(* IEC 61131-3 sources: 2026_Projet_YGO_ExcavatriceDragage/CODE_BACKUP/CODE_20260904_AvantWeekendBackup_v0.6.34/J_SUPERVISION/_BRIDGES, 13 files *)

(* ---- FB_CfgPersistBridge_BucketCfg.st ---- *)
(* =======================================================================
   💾 FB_CfgPersistBridge_BucketCfg — Pont persistance pour ST_BucketCfg
   ───────────────────────────────────────────────────────────────
   🎯 Rôle : Restauration et synchronisation bidirectionnelle IHM / Persist
   💾 Persistance : Transfert GVL_PERSISTENT <-> GVL_IHM sur Initialized
   📄 Doc métier : DOC/AF/AF_Partie-03_Contrats_Composants_v2.3.md §3
   ======================================================================= *)
FUNCTION_BLOCK FB_CfgPersistBridge_BucketCfg
VAR_OUTPUT
    // === ETATS RESTAURATION ===
    JustRestored            : BOOL;               // <-- [STAT] Vrai sur le cycle de restauration initiale
END_VAR
VAR_IN_OUT
    // === BUS CONFIGURATION ET PERSISTANCE ===
    Hmi                     : ST_BucketCfg;       // <-> [BUS] Structure de configuration IHM
    Persist                 : ST_BucketCfg;       // <-> [BUS] Structure de configuration persistante
END_VAR

JustRestored := FALSE;
IF NOT Hmi.Initialized THEN
    Hmi := Persist;
    Hmi.Initialized := TRUE;
    JustRestored := TRUE;
ELSE
    Persist := Hmi;
END_IF;

(* ---- FB_CfgPersistBridge_CommunCfg.st ---- *)
(* =======================================================================
   💾 FB_CfgPersistBridge_CommunCfg — Pont persistance pour ST_CommunCfg
   ───────────────────────────────────────────────────────────────
   🎯 Rôle : Restauration et synchronisation bidirectionnelle IHM / Persist
   💾 Persistance : Transfert GVL_PERSISTENT <-> GVL_IHM sur Initialized
   📄 Doc métier : DOC/AF/AF_Partie-03_Contrats_Composants_v2.3.md §3
   ======================================================================= *)
FUNCTION_BLOCK FB_CfgPersistBridge_CommunCfg
VAR_OUTPUT
    // === ETATS RESTAURATION ===
    JustRestored            : BOOL;               // <-- [STAT] Vrai sur le cycle de restauration initiale
END_VAR
VAR_IN_OUT
    // === BUS CONFIGURATION ET PERSISTANCE ===
    Hmi                     : ST_CommunCfg;       // <-> [BUS] Structure de configuration IHM
    Persist                 : ST_CommunCfg;       // <-> [BUS] Structure de configuration persistante
END_VAR

JustRestored := FALSE;
IF NOT Hmi.Initialized THEN
    Hmi := Persist;
    Hmi.Initialized := TRUE;
    JustRestored := TRUE;
ELSE
    Persist := Hmi;
END_IF;

(* ---- FB_CfgPersistBridge_CycleAssistToggles.st ---- *)
(* =======================================================================
   💾 FB_CfgPersistBridge_CycleAssistToggles — Pont persistance toggles assistance
   ───────────────────────────────────────────────────────────────
   🎯 Rôle : Restauration et synchronisation bidirectionnelle IHM / Persist
   💾 Persistance : Transfert GVL_PERSISTENT <-> GVL_IHM sur Initialized
   📄 Doc métier : DOC/AF/AF_Partie-03_Contrats_Composants_v2.3.md §3
   ======================================================================= *)
FUNCTION_BLOCK FB_CfgPersistBridge_CycleAssistToggles
VAR_OUTPUT
    // === ETATS RESTAURATION ===
    JustRestored            : BOOL;               // <-- [STAT] Vrai sur le cycle de restauration initiale
END_VAR
VAR_IN_OUT
    // === BUS CONFIGURATION ET PERSISTANCE ===
    Hmi                     : ST_CycleAssistToggles; // <-> [BUS] Structure de toggles IHM
    Persist                 : ST_CycleAssistToggles; // <-> [BUS] Structure de toggles persistante
END_VAR

JustRestored := FALSE;
IF NOT Hmi.Initialized THEN
    Hmi := Persist;
    Hmi.Initialized := TRUE;
    JustRestored := TRUE;
ELSE
    Persist := Hmi;
END_IF;

(* ---- FB_CfgPersistBridge_CycleCfg.st ---- *)
(* =======================================================================
   💾 FB_CfgPersistBridge_CycleCfg — Pont persistance pour ST_CycleCfg
   ───────────────────────────────────────────────────────────────
   🎯 Rôle : Restauration et synchronisation bidirectionnelle IHM / Persist
   💾 Persistance : Transfert GVL_PERSISTENT <-> GVL_IHM sur Initialized
   📄 Doc métier : DOC/AF/AF_Partie-03_Contrats_Composants_v2.3.md §3
   ======================================================================= *)
FUNCTION_BLOCK FB_CfgPersistBridge_CycleCfg
VAR_OUTPUT
    // === ETATS RESTAURATION ===
    JustRestored            : BOOL;               // <-- [STAT] Vrai sur le cycle de restauration initiale
END_VAR
VAR_IN_OUT
    // === BUS CONFIGURATION ET PERSISTANCE ===
    Hmi                     : ST_CycleCfg;        // <-> [BUS] Structure de configuration IHM
    Persist                 : ST_CycleCfg;        // <-> [BUS] Structure de configuration persistante
END_VAR

JustRestored := FALSE;
IF NOT Hmi.Initialized THEN
    Hmi := Persist;
    Hmi.Initialized := TRUE;
    JustRestored := TRUE;
ELSE
    Persist := Hmi;
END_IF;

(* ---- FB_CfgPersistBridge_CycleDiveSearchCfg.st ---- *)
(* =======================================================================
   💾 FB_CfgPersistBridge_CycleDiveSearchCfg — Pont persistance cycle plongée
   ───────────────────────────────────────────────────────────────
   🎯 Rôle : Restauration et synchronisation bidirectionnelle IHM / Persist
   💾 Persistance : Transfert GVL_PERSISTENT <-> GVL_IHM sur Initialized
   📄 Doc métier : DOC/AF/AF_Partie-03_Contrats_Composants_v2.3.md §3
   ======================================================================= *)
FUNCTION_BLOCK FB_CfgPersistBridge_CycleDiveSearchCfg
VAR_OUTPUT
    // === ETATS RESTAURATION ===
    JustRestored            : BOOL;               // <-- [STAT] Vrai sur le cycle de restauration initiale
END_VAR
VAR_IN_OUT
    // === BUS CONFIGURATION ET PERSISTANCE ===
    Hmi                     : ST_CycleDiveSearchCfg; // <-> [BUS] Structure de configuration IHM
    Persist                 : ST_CycleDiveSearchCfg; // <-> [BUS] Structure de configuration persistante
END_VAR

JustRestored := FALSE;
IF NOT Hmi.Initialized THEN
    Hmi := Persist;
    Hmi.Initialized := TRUE;
    JustRestored := TRUE;
ELSE
    Persist := Hmi;
END_IF;

(* ---- FB_CfgPersistBridge_CycleDumpAtTremieCfg.st ---- *)
(* =======================================================================
   💾 FB_CfgPersistBridge_CycleDumpAtTremieCfg — Pont persistance cycle vidage trémie
   ───────────────────────────────────────────────────────────────
   🎯 Rôle : Restauration et synchronisation bidirectionnelle IHM / Persist
   💾 Persistance : Transfert GVL_PERSISTENT <-> GVL_IHM sur Initialized
   📄 Doc métier : DOC/AF/AF_Partie-03_Contrats_Composants_v2.3.md §3
   ======================================================================= *)
FUNCTION_BLOCK FB_CfgPersistBridge_CycleDumpAtTremieCfg
VAR_OUTPUT
    // === ETATS RESTAURATION ===
    JustRestored            : BOOL;               // <-- [STAT] Vrai sur le cycle de restauration initiale
END_VAR
VAR_IN_OUT
    // === BUS CONFIGURATION ET PERSISTANCE ===
    Hmi                     : ST_CycleDumpAtTremieCfg; // <-> [BUS] Structure de configuration IHM
    Persist                 : ST_CycleDumpAtTremieCfg; // <-> [BUS] Structure de configuration persistante
END_VAR

JustRestored := FALSE;
IF NOT Hmi.Initialized THEN
    Hmi := Persist;
    Hmi.Initialized := TRUE;
    JustRestored := TRUE;
ELSE
    Persist := Hmi;
END_IF;

(* ---- FB_CfgPersistBridge_CycleExtractionCfg.st ---- *)
(* =======================================================================
   💾 FB_CfgPersistBridge_CycleExtractionCfg — Pont persistance cycle extraction
   ───────────────────────────────────────────────────────────────
   🎯 Rôle : Restauration et synchronisation bidirectionnelle IHM / Persist
   💾 Persistance : Transfert GVL_PERSISTENT <-> GVL_IHM sur Initialized
   📄 Doc métier : DOC/AF/AF_Partie-03_Contrats_Composants_v2.3.md §3
   ======================================================================= *)
FUNCTION_BLOCK FB_CfgPersistBridge_CycleExtractionCfg
VAR_OUTPUT
    // === ETATS RESTAURATION ===
    JustRestored            : BOOL;               // <-- [STAT] Vrai sur le cycle de restauration initiale
END_VAR
VAR_IN_OUT
    // === BUS CONFIGURATION ET PERSISTANCE ===
    Hmi                     : ST_CycleExtractionCfg; // <-> [BUS] Structure de configuration IHM
    Persist                 : ST_CycleExtractionCfg; // <-> [BUS] Structure de configuration persistante
END_VAR

JustRestored := FALSE;
IF NOT Hmi.Initialized THEN
    Hmi := Persist;
    Hmi.Initialized := TRUE;
    JustRestored := TRUE;
ELSE
    Persist := Hmi;
END_IF;

(* ---- FB_CfgPersistBridge_CycleMachineHomingCfg.st ---- *)
(* =======================================================================
   💾 FB_CfgPersistBridge_CycleMachineHomingCfg — Pont persistance pour ST_CycleMachineHomingCfg
   ───────────────────────────────────────────────────────────────
   🎯 Rôle : Restauration et synchronisation bidirectionnelle IHM / Persist
   💾 Persistance : Transfert GVL_PERSISTENT <-> GVL_IHM sur Initialized
   📄 Doc métier : DOC/AF/AF_Partie-03_Contrats_Composants_v2.3.md §3
   ======================================================================= *)
FUNCTION_BLOCK FB_CfgPersistBridge_CycleMachineHomingCfg
VAR_OUTPUT
    // === ETATS RESTAURATION ===
    JustRestored            : BOOL;                     // <-- [STAT] Vrai sur le cycle de restauration initiale
END_VAR
VAR_IN_OUT
    // === BUS CONFIGURATION ET PERSISTANCE ===
    Hmi                     : ST_CycleMachineHomingCfg;      // <-> [BUS] Structure de configuration IHM
    Persist                 : ST_CycleMachineHomingCfg;      // <-> [BUS] Structure de configuration persistante
END_VAR

JustRestored := FALSE;
IF NOT Hmi.Initialized THEN
    Hmi := Persist;
    Hmi.Initialized := TRUE;
    JustRestored := TRUE;
ELSE
    Persist := Hmi;
END_IF;

(* ---- FB_CfgPersistBridge_fbEncoder_Cfg.st ---- *)
(* =======================================================================
   💾 FB_CfgPersistBridge_fbEncoder_Cfg — Pont persistance pour ST_fbEncoder_Cfg
   ───────────────────────────────────────────────────────────────────────
   🎯 Rôle : restauration et synchronisation bidirectionnelle IHM / Persist.
   💾 Persistance : transfert GVL_PERSISTENT <-> GVL_IHM sur Initialized.
   📄 Doc : DOC/AF/AF_Partie-09_Fonction_Encoder_v2.4.md
   ======================================================================= *)
FUNCTION_BLOCK FB_CfgPersistBridge_fbEncoder_Cfg
VAR_OUTPUT
    // === ETATS RESTAURATION ===
    JustRestored : BOOL; // <-- [STAT] Vrai sur le cycle de restauration initiale
END_VAR
VAR_IN_OUT
    // === BUS CONFIGURATION ET PERSISTANCE ===
    Hmi    : ST_fbEncoder_Cfg; // <-> [BUS] Structure de configuration IHM commune
    Persist : ST_fbEncoder_Cfg; // <-> [BUS] Structure de configuration persistante
END_VAR

JustRestored := FALSE;
IF NOT Hmi.Initialized THEN
    Hmi := Persist;
    Hmi.Initialized := TRUE;
    JustRestored := TRUE;
ELSE
    Persist := Hmi;
END_IF;

(* ---- FB_CfgPersistBridge_fbJoystick_Cfg.st ---- *)
(* =======================================================================
   💾 FB_CfgPersistBridge_fbJoystick_Cfg — Pont persistance pour ST_fbJoystick_Cfg
   ───────────────────────────────────────────────────────────────
   🎯 Rôle : Restauration et synchronisation bidirectionnelle IHM / Persist
   💾 Persistance : Transfert GVL_PERSISTENT <-> GVL_IHM sur Initialized
   📄 Doc métier : DOC/AF/AF_Partie-08_Fonction_Joystick_v2.5.md
   ======================================================================= *)
FUNCTION_BLOCK FB_CfgPersistBridge_fbJoystick_Cfg
VAR_OUTPUT
    // === ETATS RESTAURATION ===
    JustRestored            : BOOL;                  // <-- [STAT] Vrai sur le cycle de restauration initiale
END_VAR
VAR_IN_OUT
    // === BUS CONFIGURATION ET PERSISTANCE ===
    Hmi                     : ST_fbJoystick_Cfg;     // <-> [BUS] Structure de configuration IHM
    Persist                 : ST_fbJoystick_Cfg;     // <-> [BUS] Structure de configuration persistante
END_VAR

JustRestored := FALSE;
IF NOT Hmi.Initialized THEN
    Hmi := Persist;
    Hmi.Initialized := TRUE;
    JustRestored := TRUE;
ELSE
    Persist := Hmi;
END_IF;

(* ---- FB_CfgPersistBridge_SyncCfg.st ---- *)
(* =======================================================================
   💾 FB_CfgPersistBridge_SyncCfg — Pont persistance pour ST_SyncCfg
   ───────────────────────────────────────────────────────────────
   🎯 Rôle : Restauration et synchronisation bidirectionnelle IHM / Persist
   💾 Persistance : Transfert GVL_PERSISTENT <-> GVL_IHM sur Initialized
   📄 Doc métier : DOC/AF/AF_Partie-03_Contrats_Composants_v2.3.md §3
   ======================================================================= *)
FUNCTION_BLOCK FB_CfgPersistBridge_SyncCfg
VAR_OUTPUT
    // === ETATS RESTAURATION ===
    JustRestored            : BOOL;               // <-- [STAT] Vrai sur le cycle de restauration initiale
END_VAR
VAR_IN_OUT
    // === BUS CONFIGURATION ET PERSISTANCE ===
    Hmi                     : ST_SyncCfg;         // <-> [BUS] Structure de configuration IHM
    Persist                 : ST_SyncCfg;         // <-> [BUS] Structure de configuration persistante
END_VAR

JustRestored := FALSE;
IF NOT Hmi.Initialized THEN
    Hmi := Persist;
    Hmi.Initialized := TRUE;
    JustRestored := TRUE;
ELSE
    Persist := Hmi;
END_IF;

(* ---- FB_CfgPersistBridge_TranslationCfg.st ---- *)
(* =======================================================================
   💾 FB_CfgPersistBridge_TranslationCfg — Pont persistance pour ST_TranslationCfg
   ───────────────────────────────────────────────────────────────
   🎯 Rôle : Restauration et synchronisation bidirectionnelle IHM / Persist
   💾 Persistance : Transfert GVL_PERSISTENT <-> GVL_IHM sur Initialized
   📄 Doc métier : DOC/AF/AF_Partie-11_Fonction_Translation_v2.3.md
   ======================================================================= *)
FUNCTION_BLOCK FB_CfgPersistBridge_TranslationCfg
VAR_OUTPUT
    // === ETATS RESTAURATION ===
    JustRestored            : BOOL;               // <-- [STAT] Vrai sur le cycle de restauration initiale
END_VAR
VAR_IN_OUT
    // === BUS CONFIGURATION ET PERSISTANCE ===
    Hmi                     : ST_TranslationCfg;  // <-> [BUS] Structure de configuration IHM
    Persist                 : ST_TranslationCfg;  // <-> [BUS] Structure de configuration persistante
END_VAR

JustRestored := FALSE;
IF NOT Hmi.Initialized THEN
    Hmi := Persist;
    Hmi.Initialized := TRUE;
    JustRestored := TRUE;
ELSE
    Persist := Hmi;
END_IF;

(* ---- FB_CfgPersistBridge_WinchCfg.st ---- *)
(* =======================================================================
   💾 FB_CfgPersistBridge_WinchCfg — Pont persistance pour ST_WinchCfg
   ───────────────────────────────────────────────────────────────
   🎯 Rôle : Restauration et synchronisation bidirectionnelle IHM / Persist
   💾 Persistance : Transfert GVL_PERSISTENT <-> GVL_IHM sur Initialized
   📄 Doc métier : DOC/AF/AF_Partie-10_Fonction_Winch_v2.1.md
   ======================================================================= *)
FUNCTION_BLOCK FB_CfgPersistBridge_WinchCfg
VAR_OUTPUT
    // === ETATS RESTAURATION ===
    JustRestored            : BOOL;               // <-- [STAT] Vrai sur le cycle de restauration initiale
END_VAR
VAR_IN_OUT
    // === BUS CONFIGURATION ET PERSISTANCE ===
    Hmi                     : ST_WinchCfg;        // <-> [BUS] Structure de configuration IHM
    Persist                 : ST_WinchCfg;        // <-> [BUS] Structure de configuration persistante
END_VAR

JustRestored := FALSE;
IF NOT Hmi.Initialized THEN
    Hmi := Persist;
    Hmi.Initialized := TRUE;
    JustRestored := TRUE;
ELSE
    Persist := Hmi;
END_IF;
